// TwinCAT 3 PLC project DemoLib
// Title: DemoLib
// Company: Demo
// Author: TwinCAT Explorer
// ProjectVersion: 1.0.0.0
// ProgramVersion: 3.1.4026.27
// libraries:
//   Tc2_Standard, * (Beckhoff Automation GmbH)
//   Tc2_System, * (Beckhoff Automation GmbH)
// project tree:
//   DUTs/ E_ValveState.TcDUT, ST_ValveStatus.TcDUT, T_Percent.TcDUT, U_Word.TcDUT
//   GVLs/ GVL_DemoLib.TcGVL
//   POUs/ F_Clamp.TcPOU
//   POUs/Valves/ FB_ValveBase.TcPOU, I_Valve.TcIO
// (motion and I/O tree: see PLC project machine)
// real-time tasks:
//   TASK PlcTask: cycle T#10ms, priority 20, ADS port 350
// variable links:

// ---- DUTs/E_ValveState.TcDUT
{attribute 'qualified_only'}
{attribute 'strict'}
TYPE E_ValveState :
(
	Closed := 0,
	Opening,
	Open,
	Closing,
	Error := 99
);
END_TYPE

// ---- DUTs/ST_ValveStatus.TcDUT
TYPE ST_ValveStatus :
STRUCT
	eState		: E_ValveState;
	bInterlocked	: BOOL;
	nCycles		: UDINT;
	fOpenTime	: LREAL; // s
END_STRUCT
END_TYPE

// ---- DUTs/T_Percent.TcDUT
TYPE T_Percent : LREAL;
END_TYPE

// ---- DUTs/U_Word.TcDUT
TYPE U_Word :
UNION
	nValue	: WORD;
	aBytes	: ARRAY[0..1] OF BYTE;
END_UNION
END_TYPE

// ---- GVLs/GVL_DemoLib.TcGVL
{attribute 'qualified_only'}
VAR_GLOBAL CONSTANT
	MAX_VALVES		: INT := 8;
	DEFAULT_TIMEOUT	: TIME := T#5S;
END_VAR

// ---- POUs/Valves/I_Valve.TcIO
INTERFACE I_Valve

METHOD Close : BOOL
END_METHOD

METHOD Open : BOOL
VAR_INPUT
	bForce	: BOOL;
END_VAR
END_METHOD

PROPERTY State : E_ValveState
GET // PUBLIC
END_GET
END_PROPERTY

END_INTERFACE

// ---- POUs/F_Clamp.TcPOU
FUNCTION F_Clamp : LREAL
VAR_INPUT
	fValue	: LREAL;
	fMin	: LREAL;
	fMax	: LREAL;
END_VAR

F_Clamp := MIN(MAX(fValue, fMin), fMax);

END_FUNCTION

// ---- POUs/Valves/FB_ValveBase.TcPOU
FUNCTION_BLOCK ABSTRACT FB_ValveBase IMPLEMENTS I_Valve
VAR_INPUT
	bInterlock	: BOOL;
END_VAR
VAR_OUTPUT
	stStatus	: ST_ValveStatus;
END_VAR
VAR
	tonTimeout	: TON;
END_VAR

tonTimeout(IN := stStatus.eState = E_ValveState.Opening OR stStatus.eState = E_ValveState.Closing, PT := GVL_DemoLib.DEFAULT_TIMEOUT);
IF tonTimeout.Q THEN
	stStatus.eState := E_ValveState.Error;
END_IF
stStatus.bInterlocked := bInterlock;

METHOD Close : BOOL
stStatus.eState := E_ValveState.Closing;
Close := TRUE;
END_METHOD

METHOD Open : BOOL
VAR_INPUT
	bForce	: BOOL;
END_VAR
IF bInterlock AND NOT bForce THEN
	RETURN;
END_IF
stStatus.eState := E_ValveState.Opening;
stStatus.nCycles := stStatus.nCycles + 1;
Open := TRUE;
END_METHOD

PROPERTY State : E_ValveState
GET // PUBLIC
State := stStatus.eState;
END_GET
END_PROPERTY

END_FUNCTION_BLOCK
